(* CODESYS project Overview.export

Project tree, tasks and I/O mapping:
  visualisation Overview
*)

// /Overview
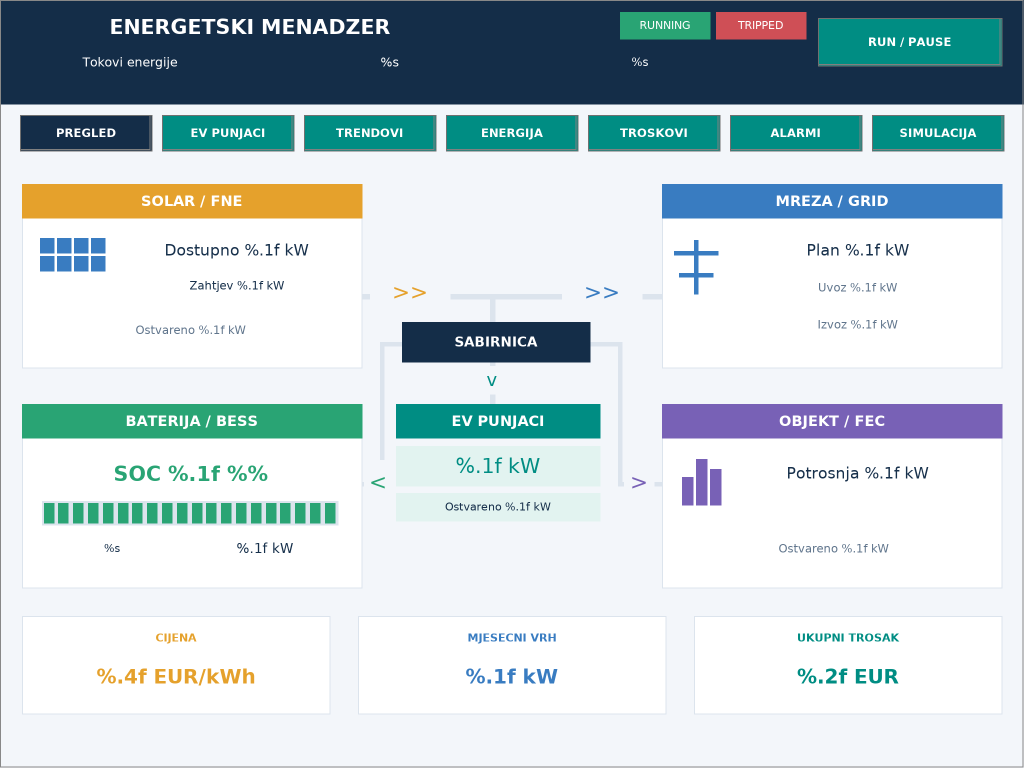
VISUALIZATION Overview  // 1024x768
    Rectangle (0,0 1024x768)
    Rectangle (0,0 1024x104)
    Rectangle (20,10 460x34), "ENERGETSKI MENADZER"
    Rectangle (20,48 220x28), "Tokovi energije"
    Rectangle (260,49 260x26), "%s", text variable: Team_HMI.sDateTime
    Rectangle (530,49 220x26), "%s", text variable: Team_HMI.sPriceMode
    Button (818,18 184x48), "RUN / PAUSE"
        toggle SimCtrl.run
    Rectangle (620,12 90x27), "PAUSED", invisible if: SimCtrl.run
    Rectangle (620,12 90x27), "RUNNING", invisible if: NOT SimCtrl.run
    Rectangle (716,12 90x27), "TRIPPED", invisible if: NOT SimCtrl.tripped
    Button (20,115 132x36), "PREGLED"
        OnMouseClick:  Assign=Overview, Type=Assignment
    Button (162,115 132x36), "EV PUNJACI"
        OnMouseClick:  Assign=EVs, Type=Assignment
    Button (304,115 132x36), "TRENDOVI"
        OnMouseClick:  Assign=Trends, Type=Assignment
    Button (446,115 132x36), "ENERGIJA"
        OnMouseClick:  Assign=Energy, Type=Assignment
    Button (588,115 132x36), "TROSKOVI"
        OnMouseClick:  Assign=Costs, Type=Assignment
    Button (730,115 132x36), "ALARMI"
        OnMouseClick:  Assign=Alarms, Type=Assignment
    Button (872,115 132x36), "SIMULACIJA"
        OnMouseClick:  Assign=Controls, Type=Assignment
    Rectangle (324,294 338x5)
    Rectangle (490,294 5x110)
    Rectangle (380,342 4x142)
    Rectangle (362,482 22x4)
    Rectangle (380,342 22x4)
    Rectangle (618,342 4x142)
    Rectangle (618,482 44x4)
    Rectangle (590,342 32x4)
    Rectangle (22,184 340x184)
    Rectangle (22,184 340x34), "SOLAR / FNE"
    Rectangle (662,184 340x184)
    Rectangle (662,184 340x34), "MREZA / GRID"
    Rectangle (22,404 340x184)
    Rectangle (22,404 340x34), "BATERIJA / BESS"
    Rectangle (662,404 340x184)
    Rectangle (662,404 340x34), "OBJEKT / FEC"
    Rectangle (40,238 14x15)
    Rectangle (57,238 14x15)
    Rectangle (74,238 14x15)
    Rectangle (91,238 14x15)
    Rectangle (40,256 14x15)
    Rectangle (57,256 14x15)
    Rectangle (74,256 14x15)
    Rectangle (91,256 14x15)
    Rectangle (128,232 218x36), "Dostupno %.1f kW", text variable: Team_HMI.rFneAvail
    Rectangle (128,271 218x29), "Zahtjev %.1f kW", text variable: Team_HMI.rFneExpected
    Rectangle (40,315 302x30), "Ostvareno %.1f kW", text variable: Team_HMI.rFneAct
    Rectangle (694,240 4x54)
    Rectangle (674,251 44x4)
    Rectangle (679,273 34x4)
    Rectangle (730,232 256x36), "Plan %.1f kW", text variable: Team_HMI.rGridPred
    Rectangle (730,273 256x29), "Uvoz %.1f kW", text variable: Team_HMI.rImportAct
    Rectangle (730,310 256x29), "Izvoz %.1f kW", text variable: Team_HMI.rExportAct
    Rectangle (370,270 80x44), ">>", invisible if: Team_HMI.rFneExpected <= 0.1
    Rectangle (562,270 80x44), "<<", invisible if: Team_HMI.rGridPred <= 0.1
    Rectangle (562,270 80x44), ">>", invisible if: Team_HMI.rGridPred >= -0.1
    Rectangle (402,322 188x40), "SABIRNICA"
    Rectangle (40,454 302x40), "SOC %.1f %%", text variable: Team_HMI.rSoc
    Rectangle (42,501 296x24)
    Rectangle (44,503 10x20), invisible if: (Team_HMI.rSoc) < 5.000
    Rectangle (58,503 10x20), invisible if: (Team_HMI.rSoc) < 10.000
    Rectangle (73,503 10x20), invisible if: (Team_HMI.rSoc) < 15.000
    Rectangle (88,503 10x20), invisible if: (Team_HMI.rSoc) < 20.000
    Rectangle (103,503 10x20), invisible if: (Team_HMI.rSoc) < 25.000
    Rectangle (118,503 10x20), invisible if: (Team_HMI.rSoc) < 30.000
    Rectangle (132,503 10x20), invisible if: (Team_HMI.rSoc) < 35.000
    Rectangle (147,503 10x20), invisible if: (Team_HMI.rSoc) < 40.000
    Rectangle (162,503 10x20), invisible if: (Team_HMI.rSoc) < 45.000
    Rectangle (177,503 10x20), invisible if: (Team_HMI.rSoc) < 50.000
    Rectangle (192,503 10x20), invisible if: (Team_HMI.rSoc) < 55.000
    Rectangle (206,503 10x20), invisible if: (Team_HMI.rSoc) < 60.000
    Rectangle (221,503 10x20), invisible if: (Team_HMI.rSoc) < 65.000
    Rectangle (236,503 10x20), invisible if: (Team_HMI.rSoc) < 70.000
    Rectangle (251,503 10x20), invisible if: (Team_HMI.rSoc) < 75.000
    Rectangle (266,503 10x20), invisible if: (Team_HMI.rSoc) < 80.000
    Rectangle (280,503 10x20), invisible if: (Team_HMI.rSoc) < 85.000
    Rectangle (295,503 10x20), invisible if: (Team_HMI.rSoc) < 90.000
    Rectangle (310,503 10x20), invisible if: (Team_HMI.rSoc) < 95.000
    Rectangle (325,503 10x20), invisible if: (Team_HMI.rSoc) < 100.000
    Rectangle (40,535 144x27), "%s", text variable: Team_HMI.sBessDir
    Rectangle (188,535 154x27), "%.1f kW", text variable: Team_HMI.rBessReq
    Rectangle (364,460 28x44), ">", invisible if: Team_HMI.rBessReq <= 0.1
    Rectangle (364,460 28x44), "<", invisible if: Team_HMI.rBessReq >= -0.1
    Rectangle (682,477 11x28)
    Rectangle (696,459 11x46)
    Rectangle (710,469 11x36)
    Rectangle (730,454 256x38), "Potrosnja %.1f kW", text variable: Team_HMI.rFec
    Rectangle (682,535 304x27), "Ostvareno %.1f kW", text variable: Team_HMI.rFecPrev
    Rectangle (624,460 30x44), ">", invisible if: Team_HMI.rFec <= 0.1
    Rectangle (396,404 204x34), "EV PUNJACI"
    Rectangle (396,446 204x40), "%.1f kW", text variable: Team_HMI.rEvReqSum
    Rectangle (396,493 204x28), "Ostvareno %.1f kW", text variable: Team_HMI.rEvActSum
    Rectangle (469,366 46x28), "v", invisible if: Team_HMI.rEvReqSum <= 0.1
    Rectangle (22,616 308x98)
    Rectangle (34,626 284x24), "CIJENA"
    Rectangle (34,657 284x39), "%.4f EUR/kWh", text variable: Team_HMI.rPrice
    Rectangle (358,616 308x98)
    Rectangle (370,626 284x24), "MJESECNI VRH"
    Rectangle (370,657 284x39), "%.1f kW", text variable: Team_HMI.rPeakMonth
    Rectangle (694,616 308x98)
    Rectangle (706,626 284x24), "UKUPNI TROSAK"
    Rectangle (706,657 284x39), "%.2f EUR", text variable: Team_Results.cost_total
END_VISUALIZATION
